(* IEC 61131-3 sources: kns-pump-station/tests/POUs/Log/FB_DeviceAudit_Test, 5 files *)

(* ---- FB_DeviceAudit_Test.decl.st ---- *)
// Назначение: набор coUnit для FB_DeviceAudit — первый вызов без событий, смена режима устройства — событие
//             101018 со значением dev_no · 10 + режим, без журнала — без ошибок. Устройства — PL.FB_DigitalInput,
//             журнал — FB_EventLog (VAR_INST), время — PL.FB_FakeTime.
// Автор:      kr0nsch
// Версия:     0.1.0
// Документ:   docs/DESIGN.md, разделы 9.3, 14.1
FUNCTION_BLOCK FB_DeviceAudit_Test EXTENDS coUnit.FB_TestSuite
VAR CONSTANT
    R_EPS : REAL := 1.0E-6;         // допуск значения события
END_VAR

(* ---- AuditLogsModeChange.method.decl.st ---- *)
// Устройство dev_no 102 из Auto в Manual: событие 101018 со значением 102 · 10 + 2 = 1022; без смены — тишина
METHOD PRIVATE AuditLogsModeChange
VAR_INST
    fbLog : FB_EventLog;            // журнал
END_VAR
VAR
    fbTime : PL.FB_FakeTime;        // подменное время
    fbDut  : FB_DeviceAudit;        // проверяемый аудит
    fbDi1  : PL.FB_DigitalInput;    // устройство dev_no 101 (режим не меняется)
    fbDi2  : PL.FB_DigitalInput;    // устройство dev_no 102
    stCmd1 : PL.ST_DigitalInputCmd;
    stCmd2 : PL.ST_DigitalInputCmd;
    stCfg  : PL.ST_DigitalInputCfg;
    stRec  : ST_EventRecord;        // запись журнала
END_VAR

(* ---- LargeDevNoValueNoOverflow.method.decl.st ---- *)
// dev_no 9999 (предел контракта, API 20.1): значение события 101018 = 9999 · 10 + 2 = 99992 без переполнения
// UINT (65535)
METHOD PRIVATE LargeDevNoValueNoOverflow
VAR_INST
    fbLog : FB_EventLog;            // журнал
END_VAR
VAR
    fbTime : PL.FB_FakeTime;        // подменное время
    fbDut  : FB_DeviceAudit;        // проверяемый аудит
    fbDi   : PL.FB_DigitalInput;    // устройство dev_no 9999
    stCmd  : PL.ST_DigitalInputCmd;
    stCfg  : PL.ST_DigitalInputCfg;
    stRec  : ST_EventRecord;        // запись журнала
END_VAR

(* ---- NoEventOnFirstCall.method.decl.st ---- *)
// Первый вызов запоминает режимы устройств без событий (режимы после старта ПЛК — из retain)
METHOD PRIVATE NoEventOnFirstCall
VAR_INST
    fbLog : FB_EventLog;            // журнал
END_VAR
VAR
    fbTime : PL.FB_FakeTime;        // подменное время
    fbDut  : FB_DeviceAudit;        // проверяемый аудит
    fbDi   : PL.FB_DigitalInput;    // устройство
    stCmd  : PL.ST_DigitalInputCmd;
    stCfg  : PL.ST_DigitalInputCfg;
END_VAR

(* ---- NoSinkIsSafe.method.decl.st ---- *)
// Без журнала (itfEvents = 0) смена режима считается, но ничего не пишется и ошибок нет
METHOD PRIVATE NoSinkIsSafe
VAR
    fbTime : PL.FB_FakeTime;        // подменное время
    fbDut  : FB_DeviceAudit;        // проверяемый аудит
    fbDi   : PL.FB_DigitalInput;    // устройство
    stCmd  : PL.ST_DigitalInputCmd;
    stCfg  : PL.ST_DigitalInputCfg;
END_VAR
